FUNCTION_BLOCK TONR //Retentive Timer
VAR_INPUT
    IN : BOOL;         // Input signal
	ResetTime: BOOL;	//Reset Accumulating Time
    PT : TIME := T#0S; // Preset time
END_VAR
VAR_OUTPUT
    Q : BOOL;          // Output signal (true when time is reached)
    ET : TIME;         // Elapsed time
END_VAR
VAR
    StartTime : TIME := T#0S; // Start time storage
    IsTiming : BOOL := FALSE; // Timing state
END_VAR

// Start or continue timing when the input is true
IF IN THEN
    IF NOT IsTiming THEN
        StartTime := DT_TO_TIME(dtRealTime) - ET; // Adjust start time if resuming
        IsTiming := TRUE;
    END_IF
    ET := DT_TO_TIME(dtRealTime) - StartTime; // Calculate elapsed time
ELSE
    IsTiming := FALSE; // Stop timing but retain elapsed time
END_IF

IF ResetTime THEN
	ResetTime:=FALSE;
	IsTiming := FALSE; // Stop timing but retain elapsed time
	ET:=T#0s;
END_IF
 
// Check if the elapsed time has reached the preset time
IF ET >= PT THEN
    Q := TRUE;
ELSE
    Q := FALSE;
END_IF

END_FUNCTION_BLOCK

(* stored: Version 1.1.0.1, ProductVersion 3.1.4024.13
   POU TONR: Id {9547d203-9a95-4810-86d6-cc5974a97350}, SpecialFunc None *)
